// Registre d'objets d'une station ou de la machine (docs/04 § 9), rempli par FB_ObjectFactory
INTERFACE I_ObjectHost

METHOD ClearObjects
END_METHOD

METHOD SetObject
VAR_INPUT
    nLocalId : UINT;
    ipObj : I_Object;
END_VAR
END_METHOD

END_INTERFACE

(* stored: Version 1.1.0.1, ProductVersion 3.1.4024.12
   Itf I_ObjectHost: Id {cefa9e00-a8e4-54fa-965f-9583d78e9364}
   Method ClearObjects: Id {9406d252-8b99-581d-8dfd-ba79230f9c9b}
   Method SetObject: Id {63477ae5-4f9f-5517-b7aa-9b2eaf5ae7a8} *)
